RoboDK station: Torre_hanoi.rdk

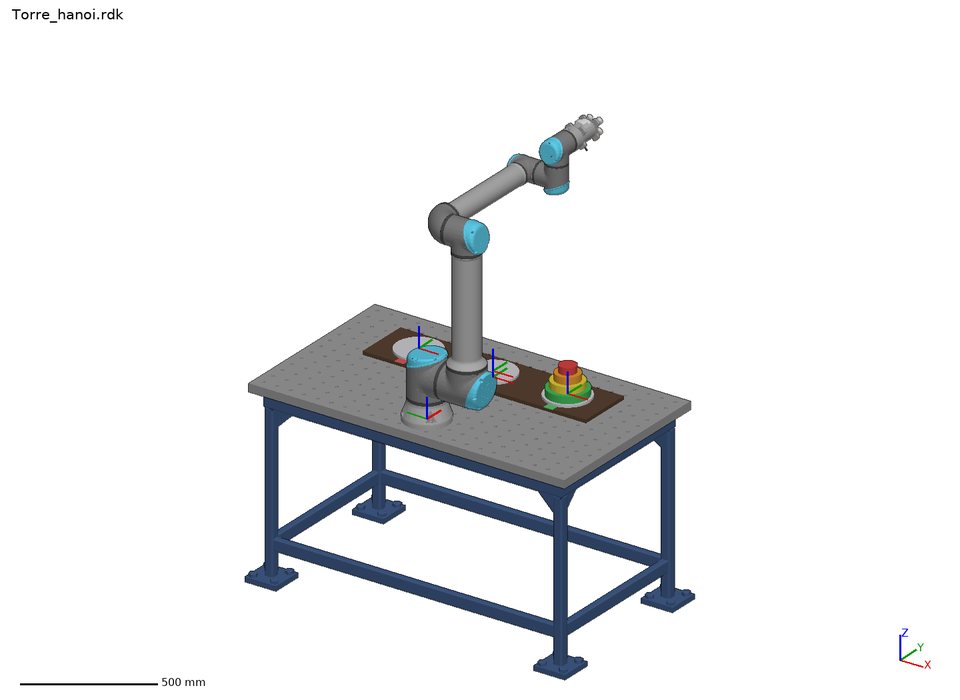
[picture v0: the station drawn from its stored meshes, robots at their saved joint values, targets as dots, program paths as lines]
Station Torre hanoi (saved by RoboDK 6.1.1). Poses are relative to the parent item; angles as X-Y-Z fixed-axis rotations.
Station parameters (name, value as stored): AltoDisco, 30, NumDiscos, 4, VelLineal, 400, VelArticular, 120, TiempoVacio, 0.3, MovimientosHechos, 15, Movimientos, 1,A,B;2,A,C;1,B,C;3,A,B;1,C,A;2,C,B;1,A,B;4,A,C;1,B,C;2,B,A;1,C,A;3,B,C;1,A,B;2,A,C;1,B,C, TotalMovimientos, 15
  - frame UR10e Base at (360, -270, 0) mm, rotated rx 0 ry 0 rz 90 deg
    - robot UR10e: 6 axes, payload 10 kg, reach 1300 mm, repeatability 0.05 mm, weight 28.9 kg
        modified DH rows (alpha deg, a mm, theta deg, d mm): 0, 0, 0, 180.7; 90, 0, 180, 0; 0, 612.6, 0, 0; 0, 571.335, 0, 174.15; -90, 0, 0, 119.85; 90, 0, 180, 116.55
        joint limits [-360, -360, -360, -360, -360, -360] to [360, 360, 360, 360, 360, 360]; home [0, -90, -90, 0, 90, 0]; saved at [0, -90, -90, 0, 90, 0]
      - tool Ventosa, TCP at (0, 0, 125) mm, size 88 x 106.8 x 127.9 mm
  - object Table 1400x800x800mm at (0, 0, 0) mm, size 1420 x 820 x 800 mm, geometry from Table-1400x800x800mm.sld
  - frame Torres at (360, 150, 0) mm
    - object Torres_base at (0, 0, 0) mm, size 990 x 240 x 15 mm, geometry from Torres_base.stl
    - frame Poste_A at (-330, 0, 25) mm
    - object Torres_apoyo_A at (-330, 0, 0) mm, size 190 x 190 x 10 mm, geometry from Torres_apoyo_A.stl
    - object Torres_letra_A at (-330, -105, 0) mm, size 40 x 40 x 2 mm, geometry from Torres_letra_A.stl
    - frame Poste_B at (0, 0, 25) mm
    - object Torres_apoyo_B at (0, 0, 0) mm, size 190 x 190 x 10 mm, geometry from Torres_apoyo_B.stl
    - object Torres_letra_B at (0, -105, 0) mm, size 40 x 40 x 2 mm, geometry from Torres_letra_B.stl
    - frame Poste_C at (330, 0, 25) mm
      - object Disco 4 at (0, 0, 0) mm, size 170 x 170 x 30 mm, geometry from Disco_4.stl
      - object Disco 3 at (0, 0, 30) mm, size 136.7 x 136.7 x 30 mm, geometry from Disco_3.stl
      - object Disco 2 at (0, 0, 60) mm, size 103.3 x 103.3 x 30 mm, geometry from Disco_2.stl
      - object Disco 1 at (0, 0, 90) mm, size 70 x 70 x 30 mm, geometry from Disco_1.stl
    - object Torres_apoyo_C at (330, 0, 0) mm, size 190 x 190 x 10 mm, geometry from Torres_apoyo_C.stl
    - object Torres_letra_C at (330, -105, 0) mm, size 40 x 40 x 2 mm, geometry from Torres_letra_C.stl
  - Python program Configurar_Parametros (listed below)
  - Python program Preparar_Torres (listed below)
  - Python program Resolver_Hanoi (listed below)
  - Python program Mover_Discos (listed below)
  - Python program Verificar_Resultado (listed below)
  - program Simulacion_Hanoi (5 instructions, listed below)

--- Python program Configurar_Parametros ---
# =====================================================================
#  Configurar_Parametros
#  Define los valores de la simulacion. Los demas programas los leen
#  como "parametros de estacion" (RDK.getParam).
# =====================================================================
from robodk.robolink import *

RDK = Robolink()

NUM_DISCOS = 4               # 3 discos = 7 movimientos, 4 = 15, 5 = 31
VEL_LINEAL = 400             # mm/s
VEL_ARTICULAR = 120          # grados/s
TIEMPO_VACIO = 0.3           # segundos para hacer o soltar el vacio de la ventosa
VEL_SIMULACION = 1           # 1 = tiempo real

RDK.setSimulationSpeed(VEL_SIMULACION)
RDK.setParam('NumDiscos', NUM_DISCOS)
RDK.setParam('VelLineal', VEL_LINEAL)
RDK.setParam('VelArticular', VEL_ARTICULAR)
RDK.setParam('TiempoVacio', TIEMPO_VACIO)
print('Parametros listos: %d discos' % NUM_DISCOS)

--- Python program Preparar_Torres ---
# =====================================================================
#  Preparar_Torres
#  Deja el juego en su estado inicial: borra los discos anteriores, apila
#  los discos nuevos en el Poste A (el mas grande abajo) y lleva el robot
#  a su posicion de reposo.
# =====================================================================
import os, math, tempfile
from robodk.robolink import *
from robodk.robomath import *

RDK = Robolink()

HOME = [0, -90, -90, 0, 90, 0]
DIAM_MIN, DIAM_MAX = 70, 170            # diametro del disco mas chico y del mas grande
COLORES = [[0.90, 0.20, 0.20], [0.95, 0.60, 0.10], [0.95, 0.85, 0.15],
           [0.20, 0.75, 0.30], [0.20, 0.45, 0.90], [0.60, 0.30, 0.80]]

N = int(float(str(RDK.getParam('NumDiscos'))))
ALTO = float(str(RDK.getParam('AltoDisco')))
poste_a = RDK.Item('Poste_A', ITEM_TYPE_FRAME)


def disco(nombre, radio, alto, rgb, padre, pose, lados=36):
    """Crea un disco (cilindro) con su origen en el centro de la base."""
    ab = [(radio * math.cos(2 * pi * k / lados), radio * math.sin(2 * pi * k / lados), 0) for k in range(lados)]
    ar = [(x, y, alto) for x, y, _ in ab]
    cb, ct = (0, 0, 0), (0, 0, alto)
    tri = []
    for k in range(lados):
        n = (k + 1) % lados
        tri += [(cb, ab[n], ab[k]), (ct, ar[k], ar[n]), (ab[k], ab[n], ar[n]), (ab[k], ar[n], ar[k])]
    ruta = os.path.join(tempfile.gettempdir(), nombre.replace(' ', '_') + '.stl')
    with open(ruta, 'w') as f:
        f.write('solid disco\n')
        for t in tri:
            f.write(' facet normal 0 0 0\n  outer loop\n')
            for v in t:
                f.write('   vertex %f %f %f\n' % v)
            f.write('  endloop\n endfacet\n')
        f.write('endsolid disco\n')
    obj = RDK.AddFile(ruta, padre)
    obj.setName(nombre)
    obj.setColor(rgb)
    obj.setPose(pose)
    return obj


for it in RDK.ItemList(ITEM_TYPE_OBJECT):
    try:
        if it.Valid() and it.Name().startswith('Disco '):
            it.Delete()
    except Exception:
        pass

# Disco N (el mas grande) abajo ... Disco 1 (el mas chico) arriba
for nivel in range(N):
    numero = N - nivel
    diam = DIAM_MIN + (DIAM_MAX - DIAM_MIN) * (numero - 1) / max(N - 1, 1)
    disco('Disco %d' % numero, diam / 2, ALTO, COLORES[(numero - 1) % len(COLORES)],
          poste_a, transl(0, 0, nivel * ALTO))

RDK.Item('UR10e', ITEM_TYPE_ROBOT).setJoints(HOME)
RDK.setParam('MovimientosHechos', 0)
print('Torres preparadas: %d discos en el Poste A' % N)

--- Python program Resolver_Hanoi ---
# =====================================================================
#  Resolver_Hanoi
#  Calcula la secuencia de movimientos con el algoritmo RECURSIVO:
#    para mover n discos de ORIGEN a DESTINO:
#      1. mover n-1 discos de ORIGEN a AUXILIAR
#      2. mover el disco n de ORIGEN a DESTINO
#      3. mover n-1 discos de AUXILIAR a DESTINO
#  La secuencia se guarda como parametro de estacion para Mover_Discos.
# =====================================================================
from robodk.robolink import *

RDK = Robolink()


def hanoi(n, origen, destino, auxiliar, movimientos):
    if n == 0:
        return
    hanoi(n - 1, origen, auxiliar, destino, movimientos)
    movimientos.append((n, origen, destino))
    hanoi(n - 1, auxiliar, destino, origen, movimientos)


N = int(float(str(RDK.getParam('NumDiscos'))))
movimientos = []
hanoi(N, 'A', 'C', 'B', movimientos)

# Formato: "disco,origen,destino;disco,origen,destino;..."
texto = ';'.join('%d,%s,%s' % m for m in movimientos)
RDK.setParam('Movimientos', texto)
RDK.setParam('TotalMovimientos', len(movimientos))

print('Secuencia calculada: %d movimientos (minimo 2^%d - 1)' % (len(movimientos), N))
for i, (d, o, de) in enumerate(movimientos, 1):
    print('  %2d. Disco %d: %s -> %s' % (i, d, o, de))

--- Python program Mover_Discos ---
# =====================================================================
#  Mover_Discos
#  El robot ejecuta la secuencia calculada por Resolver_Hanoi. En cada
#  movimiento toma el disco de ARRIBA del poste de origen con la ventosa,
#  lo sube por encima de todas las pilas, lo lleva al poste de destino y lo
#  baja justo encima del disco que ya esta ahi.
# =====================================================================
import time
from robodk.robolink import *
from robodk.robomath import *

RDK = Robolink()


def param(nombre):
    return float(str(RDK.getParam(nombre)))


robot = RDK.Item('UR10e', ITEM_TYPE_ROBOT)
tcp = RDK.Item('Ventosa', ITEM_TYPE_TOOL)
postes = {p: RDK.Item('Poste_' + p, ITEM_TYPE_FRAME) for p in 'ABC'}

HOME = [0, -90, -90, 0, 90, 0]
ALTO = param('AltoDisco')
N = int(param('NumDiscos'))
Z_SEGURA = (N + 4) * ALTO + 120         # altura de viaje: por encima de cualquier pila
ABAJO = rotx(pi)                        # ventosa mirando hacia abajo

base = robot.Parent()
robot.setPoseFrame(base)
robot.setPoseTool(tcp)
robot.setSpeed(param('VelLineal'))
robot.setSpeedJoints(param('VelArticular'))


def ir(T_mundo, lineal=True):
    T = invH(base.PoseAbs()) * T_mundo
    if lineal:
        robot.MoveL(T)
    else:
        robot.MoveJ(T)


def discos_en(poste):
    """Discos de un poste, ordenados de abajo hacia arriba."""
    d = [c for c in postes[poste].Childs() if c.Name().startswith('Disco ')]
    return sorted(d, key=lambda c: c.Pose().Pos()[2])


def sobre(poste, z):
    """Pose de la ventosa sobre el centro del poste, a la altura z (respecto al poste)."""
    return postes[poste].PoseAbs() * transl(0, 0, z) * ABAJO


def vacio(disco, padre):
    time.sleep(param('TiempoVacio') / max(RDK.SimulationSpeed(), 0.1))
    disco.setParentStatic(padre)


texto = str(RDK.getParam('Movimientos'))
movimientos = [m.split(',') for m in texto.split(';') if m]
total = len(movimientos)

robot.MoveJ(HOME)
ir(sobre('A', Z_SEGURA), lineal=False)

for i, (num, origen, destino) in enumerate(movimientos, 1):
    RDK.ShowMessage('Movimiento %d de %d: Disco %s, de %s a %s' % (i, total, num, origen, destino), False)

    # Tomar el disco de arriba del origen
    pila = discos_en(origen)
    disco = pila[-1]
    if disco.Name() != 'Disco ' + num:
        raise Exception('Se esperaba el Disco %s arriba del poste %s' % (num, origen))
    z_tapa = len(pila) * ALTO
    ir(sobre(origen, Z_SEGURA))
    ir(sobre(origen, z_tapa))
    vacio(disco, tcp)
    ir(sobre(origen, Z_SEGURA))

    # Llevarlo al destino y apoyarlo sobre la pila que hay ahi
    z_dejar = (len(discos_en(destino)) + 1) * ALTO
    ir(sobre(destino, Z_SEGURA))
    ir(sobre(destino, z_dejar))
    vacio(disco, postes[destino])
    ir(sobre(destino, Z_SEGURA))

    RDK.setParam('MovimientosHechos', i)

robot.MoveJ(HOME)
print('Secuencia completada: %d movimientos' % total)

--- Python program Verificar_Resultado ---
# =====================================================================
#  Verificar_Resultado
#  Comprueba que todos los discos terminaron en el Poste C, ordenados del
#  mas grande (abajo) al mas chico (arriba), y muestra el resultado.
# =====================================================================
from robodk.robolink import *

RDK = Robolink()

N = int(float(str(RDK.getParam('NumDiscos'))))
hechos = int(float(str(RDK.getParam('MovimientosHechos'))))
poste_c = RDK.Item('Poste_C', ITEM_TYPE_FRAME)

discos = [c for c in poste_c.Childs() if c.Name().startswith('Disco ')]
discos.sort(key=lambda c: c.Pose().Pos()[2])              # de abajo hacia arriba
numeros = [int(c.Name().split()[1]) for c in discos]

if numeros == list(range(N, 0, -1)):
    msg = 'Torre resuelta: %d discos en el Poste C en %d movimientos (minimo 2^%d - 1 = %d).' % (
        N, hechos, N, 2 ** N - 1)
else:
    msg = 'La torre NO quedo bien: en el Poste C hay %s' % numeros
RDK.ShowMessage(msg, True)
print(msg)

--- program Simulacion_Hanoi (robot UR10e) ---
  Llamar Configurar_Parametros
  Llamar Preparar_Torres
  Llamar Resolver_Hanoi
  Llamar Mover_Discos
  Llamar Verificar_Resultado
